Staubli VAL3: main.pgx

program main()
begin
  close(tCurrentTool)
  pPointRx.config.shoulder = lefty
  pPointRx.config.elbow = epositive
  pPointRx.config.wrist = wpositive
  pPointRx2.config.shoulder = lefty
  pPointRx2.config.elbow = epositive
  pPointRx2.config.wrist = wpositive
  mCurrentSpeed.tvel = 100.00
  mCurrentSpeed.blend = joint
  mCurrentSpeed.reach = 0.010
  mCurrentSpeed.leave = 0.010
  // Program MAIN_1 start
  // Program generated by RoboDK v5.6.9 for RoboDK Industrial on 26/02/2024 09:58:20
  // Using nominal kinematics.
  call MoveJoint(-0.00000,0.00000,0.00000,0.00000,0.00000,-0.00000)
  call MoveJoint(0.00000,3.21124,-15.42370,0.00000,12.21250,-0.00000)
  pPointRx.config.wrist = wnegative
  call MoveLine(1015.000,0.000,1272.000,0.000,90.000,0.000)
  Output[5]=true
  Output[5]=true
  Output[5]=0.5
  Output[5]=true
  Output[5]=true
  Output[5]=true
  Output[5]=0.5
  Output[5]=true
  var=val
  var=val
  watch(Input[5]==true)
  watch(Input[5]==true)
  watch(Input[5]==0.5)
  watch(Input[5]==true)
  watch(Input[5]==true,100.0)
  watch(var==val)
  watch(var==val,100.0)
  popUpMsg("Message")
  //call prog:REMOTE_PROG_CALL_171()
  CODE_INSERT_172
  // Insert Comment
  mCurrentSpeed.reach = 10.000
  mCurrentSpeed.leave = 10.000
  call MoveJoint(-29.33220,46.67700,-0.02452,26.54560,25.39570,-51.63400)
  mCurrentSpeed.reach = -1.000
  mCurrentSpeed.leave = -1.000
  mCurrentSpeed.tvel = 100.000
  pPointRx.config.wrist = wpositive
  call MoveLine(187.786,125.499,139.112,-179.996,0.180,179.997)
  Output[5]=true
  //call prog:PICK_PART_111()
  mCurrentSpeed.reach = 10.000
  mCurrentSpeed.leave = 10.000
  mCurrentSpeed.tvel = 300.000
  // Linear movement using joint targets is not supported. Change the target type to cartesian or use a joint movement.
  call MoveLine(187.272,447.522,305.347,179.998,0.185,-179.999)
  mCurrentSpeed.reach = -1.000
  mCurrentSpeed.leave = -1.000
  mCurrentSpeed.tvel = 100.000
  // MoveSearch command not implemented
  call MoveLine(187.851,447.517,126.235,179.998,0.185,-179.999)
  Output[5]=false
  //call prog:PLACE_PART_112()
  mCurrentSpeed.reach = 10.000
  mCurrentSpeed.leave = 10.000
  call MoveLine(187.272,447.522,305.347,179.998,0.185,-179.999)
  mCurrentSpeed.reach = 25.000
  mCurrentSpeed.leave = 25.000
  call MoveJoint(52.18600,45.67580,6.92000,66.73420,19.93230,-92.73000)
  call MoveCirc(430.047,43.774,231.503,-171.221,7.036,133.902,109.688,-153.222,161.073,-171.221,7.036,133.902)
  // Circular movement using joint targets is not supported. Change the target type to cartesian or use a joint movement.
  mCurrentSpeed.reach = -1.000
  mCurrentSpeed.leave = -1.000
  call MoveLine(312.208,292.214,255.156,-171.221,7.036,133.902)
  call MoveJoint(-0.00000,0.00000,0.00000,0.00000,0.00000,-0.00000)
  // Warning: This post processor is meant to use one reference frame. Errors might follow.
  call MoveJoint(88.67600,29.60160,-6.42883,-1.98422,49.47920,4.54769)
  call MoveLine(19.898,174.307,19.008,174.554,-0.000,94.906)
  call MoveLine(378.402,174.416,18.997,174.554,-0.000,94.906)
  call MoveLine(380.996,112.363,34.882,161.791,-0.000,95.030)
  call MoveLine(16.551,114.359,34.226,161.791,-0.000,95.030)
  call MoveLine(26.434,54.524,46.072,-175.632,0.000,95.445)
  call MoveLine(385.448,48.050,45.137,-168.767,0.000,95.484)
  call MoveLine(385.448,-1.625,295.251,-168.767,0.000,95.484)
  call MoveJoint(-0.00000,0.00000,0.00000,0.00000,0.00000,-0.00000)
  //call prog:EVENT_PROG_START_101()
  mCurrentSpeed.reach = 1.000
  mCurrentSpeed.leave = 1.000
  mCurrentSpeed.tvel = 1000.000
  // Warning: This post processor is meant to use one reference frame. Errors might follow.
  // Show Tool 1
  call MoveJoint(-68.09030,24.20190,26.78550,38.21340,36.20170,-98.79640)
  //call prog:EVENT_PATH_APPROACH_102()
  call MoveLine(-49.895,253.259,319.999,-179.647,0.025,90.000)
  call MoveLine(0.000,250.000,270.000,-179.647,0.025,90.000)
  //call prog:EVENT_PATH_START_103()
  mCurrentSpeed.tvel = 50.000
  call MoveLine(35.579,247.455,270.000,-179.655,0.075,90.000)
  call MoveLine(70.433,239.873,270.000,-179.669,0.124,89.999)
  call MoveLine(103.854,227.408,270.000,-179.690,0.169,89.999)
  call MoveLine(135.160,210.313,270.000,-179.717,0.212,89.999)
  call MoveLine(163.715,188.937,270.000,-179.750,0.250,89.999)
  call MoveLine(188.937,163.715,270.000,-179.788,0.283,89.999)
  call MoveLine(210.313,135.160,270.000,-179.830,0.311,89.999)
  call MoveLine(227.408,103.854,270.000,-179.876,0.332,89.999)
  call MoveLine(239.873,70.433,270.000,-179.925,0.346,90.000)
  call MoveLine(247.455,35.579,270.000,-179.975,0.353,90.000)
  call MoveLine(250.000,0.000,270.000,179.975,0.353,90.000)
  call MoveLine(247.455,-35.579,270.000,179.925,0.346,90.000)
  call MoveLine(239.873,-70.433,270.000,179.876,0.332,90.001)
  call MoveLine(227.408,-103.854,270.000,179.830,0.311,90.001)
  call MoveLine(210.313,-135.160,270.000,179.788,0.283,90.001)
  call MoveLine(188.937,-163.715,270.000,179.750,0.250,90.001)
  call MoveLine(163.715,-188.937,270.000,179.717,0.212,90.001)
  call MoveLine(135.160,-210.313,270.000,179.689,0.170,90.001)
  call MoveLine(103.854,-227.408,270.000,179.668,0.124,90.001)
  call MoveLine(70.433,-239.873,270.000,179.654,0.075,90.000)
  call MoveLine(35.579,-247.455,270.000,179.647,0.025,90.000)
  call MoveLine(0.000,-250.000,270.000,179.647,0.025,90.000)
  call MoveLine(0.000,-250.000,270.000,179.647,-0.025,90.000)
  call MoveLine(-35.579,-247.455,270.000,179.654,-0.075,90.000)
  call MoveLine(-70.433,-239.873,270.000,179.669,-0.124,89.999)
  call MoveLine(-103.854,-227.408,270.000,179.690,-0.169,89.999)
  call MoveLine(-135.160,-210.313,270.000,179.717,-0.212,89.999)
  call MoveLine(-163.715,-188.937,270.000,179.750,-0.250,89.999)
  call MoveLine(-188.937,-163.715,270.000,179.788,-0.283,89.999)
  call MoveLine(-210.313,-135.160,270.000,179.831,-0.310,89.999)
  call MoveLine(-227.408,-103.854,270.000,179.877,-0.331,89.999)
  call MoveLine(-239.873,-70.433,270.000,179.925,-0.346,90.000)
  call MoveLine(-247.455,-35.579,270.000,179.975,-0.353,90.000)
  call MoveLine(-250.000,0.000,270.000,-179.975,-0.353,90.000)
  call MoveLine(-247.455,35.579,270.000,-179.925,-0.345,90.000)
  call MoveLine(-239.873,70.433,270.000,-179.877,-0.331,90.001)
  call MoveLine(-227.408,103.854,270.000,-179.830,-0.311,90.001)
  call MoveLine(-210.313,135.160,270.000,-179.788,-0.283,90.001)
  call MoveLine(-188.937,163.715,270.000,-179.750,-0.250,90.001)
  call MoveLine(-163.715,188.937,270.000,-179.717,-0.212,90.001)
  call MoveLine(-135.160,210.313,270.000,-179.690,-0.169,90.001)
  call MoveLine(-103.854,227.408,270.000,-179.668,-0.124,90.001)
  call MoveLine(-70.433,239.873,270.000,-179.654,-0.075,90.000)
  call MoveLine(-35.579,247.455,270.000,-179.647,-0.025,90.000)
  call MoveLine(0.000,250.000,270.000,-179.647,-0.025,90.000)
  mCurrentSpeed.tvel = 1000.000
  //call prog:EVENT_PATH_FINISH_105()
  call MoveLine(49.895,253.258,319.999,-179.647,-0.025,90.000)
  call MoveLine(49.939,252.642,419.997,-179.647,-0.025,90.000)
  //call prog:EVENT_PATH_RETRACT_106()
  //call prog:EVENT_PROG_FINISH_107()
  // Warning: This post processor is meant to use one reference frame. Errors might follow.
  call MoveJoint(-29.33220,46.67700,-0.02452,26.54560,25.39570,-51.63400)
  delay(1.250)
  call MoveLine(187.786,125.499,139.112,-179.996,0.180,179.997)
  watch(Input[1]==true)
  call MoveLine(187.264,125.487,305.356,180.000,0.184,-180.000)
  //call prog:PROG 1 _.-[]/\;,><&*:%=+@!#^|?^ with a very long name and special characters()

  waitEndMove()
  // Program MAIN_1 end
  // Program PROG 1 _.-[]/\;,><&*:%=+@!#^|?^ with a very long name and special characters start
  // This is a subprogram call to PROG_1
  // Warning: This post processor is meant to use one reference frame. Errors might follow.
  call MoveJoint(-0.00000,0.00000,0.00000,0.00000,0.00000,-0.00000)

  waitEndMove()
  // Program PROG 1 _.-[]/\;,><&*:%=+@!#^|?^ with a very long name and special characters end

end
